FUNCTION_BLOCK StopFeed (* Basic Function Block Type *)
  (* Standard: 61499-2 *)
  (* Version 0.0, 10/5/2026, Schneider Electric, Template *)
  PACKAGE SE.Nereda;
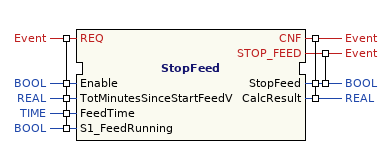
  EVENT_INPUT
    REQ WITH FeedTime, TotMinutesSinceStartFeedV, S1_FeedRunning, Enable; (* Normal Execution Request *)
  END_EVENT
  EVENT_OUTPUT
    CNF WITH StopFeed, CalcResult; (* Execution Confirmation *)
    STOP_FEED WITH StopFeed;
  END_EVENT
  VAR_INPUT
    Enable : BOOL;
    TotMinutesSinceStartFeedV : REAL; (* Input event qualifier *)
    FeedTime : TIME;
    S1_FeedRunning : BOOL;
  END_VAR
  VAR_OUTPUT
    StopFeed : BOOL; (* Output event qualifier *)
    CalcResult : REAL;
  END_VAR
  VAR
    InFeedTime : REAL;
    StopCmd : BOOL;
  END_VAR
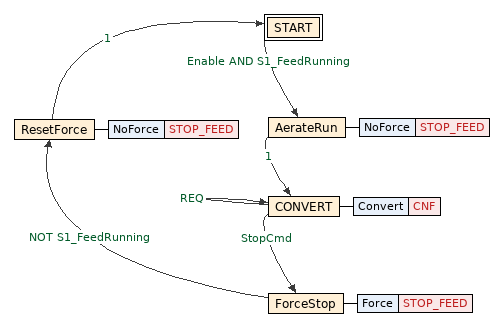
  EC_STATES
    START; (* Initial State *)
    AerateRun : NoForce -> STOP_FEED;
    ForceStop : Force -> STOP_FEED;
    ResetForce : NoForce -> STOP_FEED;
    CONVERT : Convert -> CNF;
  END_STATES
  EC_TRANSITIONS
    CONVERT TO ForceStop := StopCmd;
    ForceStop TO ResetForce := NOT S1_FeedRunning;
    AerateRun TO CONVERT := 1;
    CONVERT TO CONVERT := REQ;
    START TO AerateRun := Enable AND S1_FeedRunning;
    ResetForce TO START := 1;
  END_TRANSITIONS
  ALGORITHM NoForce IN ST:
;
StopFeed := FALSE;
  END_ALGORITHM
  ALGORITHM Convert IN ST:
;
InFeedTime := TIME_TO_REAL(FeedTime) / 60000.0;

CalcResult := InFeedTime - TotMinutesSinceStartFeedV;

StopCmd := CalcResult <= 0;
  END_ALGORITHM
  ALGORITHM Force IN ST:
;
StopFeed := TRUE;
  END_ALGORITHM
END_FUNCTION_BLOCK
